// TIA Portal V20 export
// export: Created 2026-10-19T18:03:58.3120852Z, ExportSetting WithDefaults, DisplayName Totally Integrated Automation Portal, DisplayVersion V20 Update 6, DisplayName TIA Portal Openness, DisplayVersion V20 Update 6, DisplayName TIA Portal Version Control Interface, DisplayVersion V20 Update 6, DisplayName SINAMICS Startdrive Advanced, DisplayVersion V20 SP1, DisplayName SINAMICS Startdrive G130, G150, S120, S150, SINAMICS MV, G220, S200, S210, DisplayVersion V20 SP1, DisplayName SINAMICS Startdrive G110M, G120, G120C, G120D, G120P, G115D, DisplayVersion V20 SP1, DisplayName STEP 7 Professional, DisplayVersion V20 Update 6, DisplayName STEP 7 Safety, DisplayVersion V20 Update 2, DisplayName WinCC Basic/Comfort/Advanced, DisplayVersion V20 Update 6, DisplayName WinCC Unified, DisplayVersion V20 Update 6
DATA_BLOCK "PConveyor_3_FB_DB"   // DB88
AUTHOR : Mertin Coetzee
VERSION : 0.1
// stored: AutoNumber true, DBAccessibleFromOPCUA true, DBAccessibleFromWebserver true, InstanceOfName PConveyor_3_FB, InstanceOfType FB
"PConveyor_3_FB"
   // VAR_INPUT
   //    Cnv_Settings : "PopUp_Cnv_Settings";
   //    TimeStartBoost_Chain : UInt;
   //    TimeStartBoost_Roller : UInt;
   // END_VAR
   // VAR_IN_OUT
   //    Cnv_Control : "PopUp_Cnv_Control";
   //    SinaSpeed_Roller : SinaSpeed;
   //    SinaSpeed_Chain : SinaSpeed;
   //    SinaSpeed_Lift : SinaSpeed;
   // END_VAR
   // VAR
   //    State : UInt;
   //    Timer_TC : TON_TIME;
   //    Timer_Transfer { S7_SetPoint := 'True'} : TON_TIME;
   //    Watchdog { S7_SetPoint := 'True'} : TON_TIME;
   //    Transfer_Direction { S7_SetPoint := 'True'} : String;
   //    MainSetpoint_Roller : Int;
   //    MainSetpoint_Chain : Int;
   //    MainSetpoint_Lift : Int;
   //    IEC_Timer_0_Instance_1 { S7_SetPoint := 'True'} : TON_TIME;
   //    R_TRIG_Instance { S7_SetPoint := 'True'} : R_TRIG;
   // END_VAR
BEGIN
END_DATA_BLOCK
